Fanuc KAREL source: kb00164.KL

-- PROVISIONAL review KL for V770-1; original PC SHA256 e5534e3e9f9b4815ad5a45e76811eaa719652932884757e5dc1aad792174567a
-- Incomplete behavior may be omitted. Consult companion uncertainty JSON. Do not deploy.
PROGRAM KB00164
%NOLOCKGROUP
BEGIN
  -- UNRESOLVED_PC offsets 5-12; opcodes 9D,23
  -- UNRESOLVED_PC offsets 17-24; opcodes 9D,23
  -- UNRESOLVED_PC offsets 29-51; opcodes 27,22,22,22,31
  -- UNRESOLVED_PC offsets 56-60; opcodes 7F
END KB00164
